SYSTEM System
  DEVICE EcoRT_0 : Soft_dPAC
    RESOURCE RES0 : EMB_RES_ECO
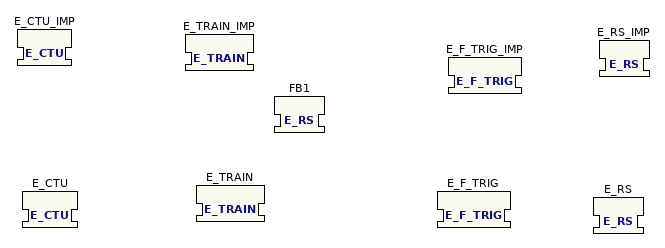
      FBS
        FB1 : E_RS;
        E_TRAIN_IMP : E_TRAIN;
        E_TRAIN : E_TRAIN;
        E_F_TRIG_IMP : E_F_TRIG;
        E_F_TRIG : E_F_TRIG;
        E_CTU_IMP : E_CTU;
        E_CTU : E_CTU;
        E_RS_IMP : E_RS;
        E_RS : E_RS;
      END_FBS
    END_RESOURCE
  END_DEVICE
END_SYSTEM
